SUBAPPLICATION RedWhiteBackground4 (* Hintergrundfarbe (TRUE -> Rot, FALSE -> Weiß) für 4 Objekte *)
  (* Standard: 61499-2 *)
  (* Version 1.0, 2026-07-21, franz, Meisterschulen am Ostbahnhof *)
  PACKAGE MyLib::sys;
  IMPORT isobus::UT::Q::const::IDs::ID_NULL;
  IMPORT isobus::UT::Q::const::colours;
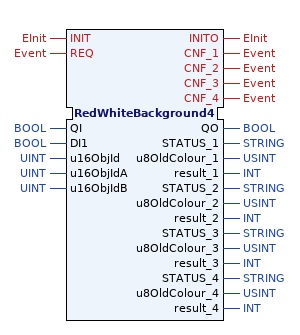
  EVENT_INPUT
    INIT : EInit; (* Initialization Request *)
    REQ; (* Normal Execution Request *)
  END_EVENT
  EVENT_OUTPUT
    INITO : EInit; (* Initialization Confirm *)
    CNF_1;
    CNF_2;
    CNF_3;
    CNF_4;
  END_EVENT
  VAR_INPUT
    QI : BOOL := TRUE; (* Quality Input - TRUE to enable service *)
    DI1 : BOOL; (* Selector *)
    u16ObjId : UINT := ID_NULL; (* Object ID Softkey *)
    u16ObjIdA : UINT := ID_NULL; (* Object ID AUX *)
    u16ObjIdB : UINT := ID_NULL; (* Object ID Button *)
  END_VAR
  VAR_OUTPUT
    QO : BOOL; (* Quality Output - TRUE if service executed successfully (AND aller Instanzen) *)
    STATUS_1 : STRING; (* Service Status *)
    u8OldColour_1 : USINT; (* Old value of ID *)
    result_1 : INT; (* retval see description *)
    STATUS_2 : STRING; (* Service Status *)
    u8OldColour_2 : USINT; (* Old value of ID *)
    result_2 : INT; (* retval see description *)
    STATUS_3 : STRING; (* Service Status *)
    u8OldColour_3 : USINT; (* Old value of ID *)
    result_3 : INT; (* retval see description *)
    STATUS_4 : STRING; (* Service Status *)
    u8OldColour_4 : USINT; (* Old value of ID *)
    result_4 : INT; (* retval see description *)
  END_VAR
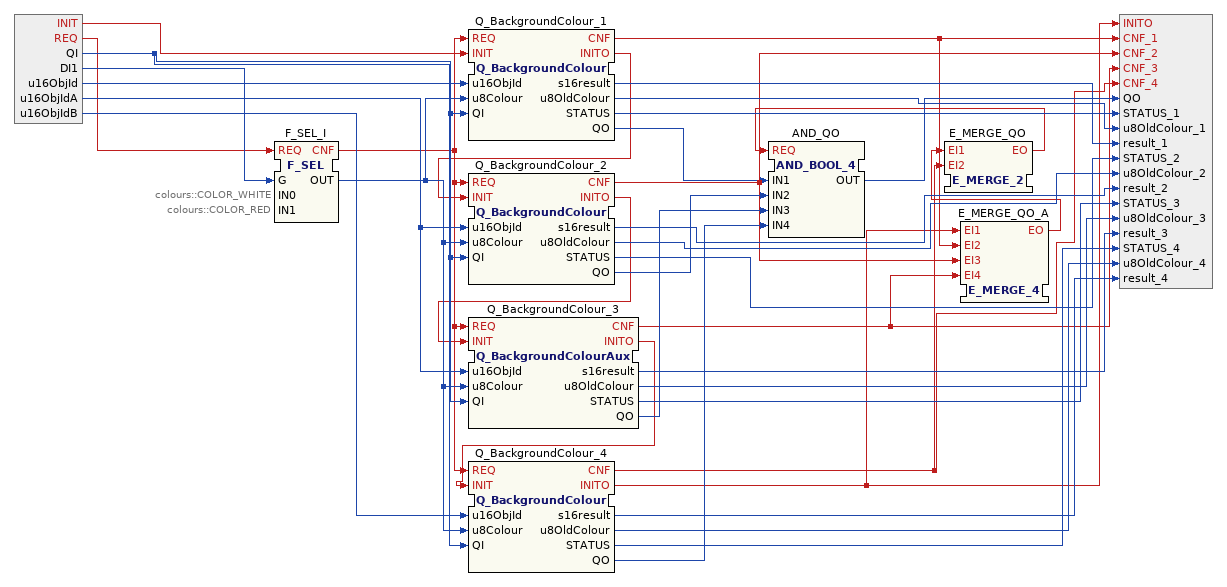
  FBS
    Q_BackgroundColour_1 : isobus::UT::Q::Q_BackgroundColour;
    Q_BackgroundColour_2 : isobus::UT::Q::Q_BackgroundColour;
    Q_BackgroundColour_3 : isobus::UT::Q::Q_BackgroundColourAux;
    Q_BackgroundColour_4 : isobus::UT::Q::Q_BackgroundColour;
    F_SEL_I : iec61131::selection::F_SEL(IN0 := colours::COLOR_WHITE, IN1 := colours::COLOR_RED);
    E_MERGE_QO_A : iec61499::events::E_MERGE_4;
    E_MERGE_QO : iec61499::events::E_MERGE_2;
    AND_QO : iec61131::booleanOperators::AND_BOOL_4;
  END_FBS
  EVENT_CONNECTIONS
    REQ TO F_SEL_I.REQ;
    Q_BackgroundColour_1.CNF TO CNF_1;
    Q_BackgroundColour_2.CNF TO CNF_2;
    Q_BackgroundColour_3.CNF TO CNF_3;
    Q_BackgroundColour_4.CNF TO CNF_4;
    F_SEL_I.CNF TO Q_BackgroundColour_1.REQ;
    F_SEL_I.CNF TO Q_BackgroundColour_4.REQ;
    F_SEL_I.CNF TO Q_BackgroundColour_3.REQ;
    F_SEL_I.CNF TO Q_BackgroundColour_2.REQ;
    INIT TO Q_BackgroundColour_1.INIT;
    Q_BackgroundColour_1.INITO TO Q_BackgroundColour_2.INIT;
    Q_BackgroundColour_2.INITO TO Q_BackgroundColour_3.INIT;
    Q_BackgroundColour_3.INITO TO Q_BackgroundColour_4.INIT;
    Q_BackgroundColour_4.INITO TO INITO;
    Q_BackgroundColour_4.INITO TO E_MERGE_QO_A.EI1;
    Q_BackgroundColour_1.CNF TO E_MERGE_QO_A.EI2;
    Q_BackgroundColour_2.CNF TO E_MERGE_QO_A.EI3;
    Q_BackgroundColour_3.CNF TO E_MERGE_QO_A.EI4;
    E_MERGE_QO_A.EO TO E_MERGE_QO.EI1;
    Q_BackgroundColour_4.CNF TO E_MERGE_QO.EI2;
    E_MERGE_QO.EO TO AND_QO.REQ;
  END_CONNECTIONS
  DATA_CONNECTIONS
    DI1 TO F_SEL_I.G;
    u16ObjId TO Q_BackgroundColour_1.u16ObjId;
    Q_BackgroundColour_1.s16result TO result_1;
    Q_BackgroundColour_1.u8OldColour TO u8OldColour_1;
    Q_BackgroundColour_1.STATUS TO STATUS_1;
    F_SEL_I.OUT TO Q_BackgroundColour_1.u8Colour;
    u16ObjIdA TO Q_BackgroundColour_2.u16ObjId;
    Q_BackgroundColour_2.s16result TO result_2;
    Q_BackgroundColour_2.u8OldColour TO u8OldColour_2;
    Q_BackgroundColour_2.STATUS TO STATUS_2;
    F_SEL_I.OUT TO Q_BackgroundColour_2.u8Colour;
    u16ObjIdA TO Q_BackgroundColour_3.u16ObjId;
    Q_BackgroundColour_3.s16result TO result_3;
    Q_BackgroundColour_3.u8OldColour TO u8OldColour_3;
    Q_BackgroundColour_3.STATUS TO STATUS_3;
    F_SEL_I.OUT TO Q_BackgroundColour_3.u8Colour;
    u16ObjIdB TO Q_BackgroundColour_4.u16ObjId;
    Q_BackgroundColour_4.s16result TO result_4;
    Q_BackgroundColour_4.u8OldColour TO u8OldColour_4;
    Q_BackgroundColour_4.STATUS TO STATUS_4;
    F_SEL_I.OUT TO Q_BackgroundColour_4.u8Colour;
    QI TO Q_BackgroundColour_1.QI;
    QI TO Q_BackgroundColour_2.QI;
    QI TO Q_BackgroundColour_3.QI;
    QI TO Q_BackgroundColour_4.QI;
    Q_BackgroundColour_1.QO TO AND_QO.IN1;
    Q_BackgroundColour_2.QO TO AND_QO.IN2;
    Q_BackgroundColour_3.QO TO AND_QO.IN3;
    Q_BackgroundColour_4.QO TO AND_QO.IN4;
    AND_QO.OUT TO QO;
  END_CONNECTIONS
END_SUBAPPLICATION
